// TIA Portal V20 export
// export: Created 2026-10-20T12:53:02.8924385Z, ExportSetting WithDefaults, DisplayName Totally Integrated Automation Portal, DisplayVersion V20 Update 6, DisplayName TIA Portal Openness, DisplayVersion V20 Update 6, DisplayName TIA Portal Version Control Interface, DisplayVersion V20 Update 6, DisplayName SINAMICS Startdrive Advanced, DisplayVersion V20 SP1, DisplayName SINAMICS Startdrive G130, G150, S120, S150, SINAMICS MV, G220, S200, S210, DisplayVersion V20 SP1, DisplayName SINAMICS Startdrive G110M, G120, G120C, G120D, G120P, G115D, DisplayVersion V20 SP1, DisplayName STEP 7 Professional, DisplayVersion V20 Update 6, DisplayName STEP 7 Safety, DisplayVersion V20 Update 2, DisplayName WinCC Basic/Comfort/Advanced, DisplayVersion V20 Update 6, DisplayName WinCC Unified, DisplayVersion V20 Update 6
FUNCTION "VTD_Status_Update_FC" : Void   // FC48, SCL
{ S7_Optimized_Access := 'TRUE' }
VERSION : 0.1
// stored: AutoNumber true, IsIECCheckEnabled false, SetENOAutomatically false, UDAEnableTagReadback false
   VAR_INPUT
      Infeed_Auto_Mode : Bool;
      Infeed_Manual_Mode : Bool;
      Infeed_Maintenance : Bool;
      Infeed_Alarm : Bool;
      Infeed_Ready : Bool;
      Outfeed_Auto_Mode : Bool;
      Pallet_ID : Array[1..100] of Byte;
   END_VAR
   VAR_OUTPUT
      SM_To_LGX_VTD_Status : Byte;
   END_VAR
   VAR_IN_OUT
      Pallet_ID_Received : Bool;
   END_VAR
   VAR_TEMP
      tStatusByte : Byte;
      ArrayHasData : Bool;
      i : UInt;
   END_VAR
BEGIN
   #tStatusByte := 0;

       #tStatusByte.%X0 := #Infeed_Auto_Mode;
       #tStatusByte.%X1 := #Infeed_Manual_Mode;
       #tStatusByte.%X2 := #Infeed_Maintenance;
       #tStatusByte.%X3 := #Infeed_Ready;
       #tStatusByte.%X4 := #Infeed_Alarm;

       #ArrayHasData := FALSE;

       FOR #i := 1 TO 100 DO
           IF #Pallet_ID[#i] <> 0 THEN
               #ArrayHasData := TRUE;
               EXIT;
           END_IF;
       END_FOR;

       #tStatusByte.%X5 := #Pallet_ID_Received AND #ArrayHasData;
       #tStatusByte.%X6 := #Outfeed_Auto_Mode;

       IF #Pallet_ID_Received AND NOT #ArrayHasData THEN
           #Pallet_ID_Received := FALSE;
       END_IF;

       // Bit 5, 6: Free
       // 
       #SM_To_LGX_VTD_Status := #tStatusByte;
END_FUNCTION
